// TIA Portal V20 export
FUNCTION "POS3_0_Teileauswertung" : Void   // FC60, STL
TITLE = Teileauswertung
{ S7_Optimized_Access := 'FALSE' }
   VAR_TEMP
      RetVal : Int;
   END_VAR
BEGIN
END_FUNCTION
